Fanuc KAREL source: KT00591.KL

PROGRAM KT00591
%NOLOCKGROUP
VAR
  S1: STRING[80]
  R2: REAL
  OUT: STRING[80]
BEGIN
  S1 = 'A'
    R2 = 3.0
  OUT = S1 + R2
END KT00591
